(* IEC 61131-3 sources: Test-Git_ESME26/TestProgettoESME_26.fbsproj/PacDriveLib Migration/Motion/Positioning, 3 files *)

(* ---- PDL_FB_EndlessFeed.fb.st ---- *)
FUNCTION_BLOCK PDL_FB_EndlessFeed

VAR_INPUT
	i_xEnable					: BOOL;			(* Enable of FB *)
	i_ifDrive					: MOIN.IF_Axis;	(* Axis *)
	i_lrVel 					: LREAL;		(* Ceiling velocity in units/sec, -MaxVel to +MaxVel *)
	i_lrAcc  					: LREAL;		(* Acceleration units/s^2, value: 0...lrLimitMaxAccDec *)
	i_lrDec 					: LREAL;		(* Deceleration units/s^2, value: 0...lrLimitMaxAccDec *)
	i_lrJerk					: LREAL;		(* Jerk units/s^3, value: >0 *)
	i_lrPeriod					: LREAL;		(* LINEAR axis: the position is kept within the period value (0 … i_lrPeriod), in units, must be > 0
												   MODULO axis: value is ignored -> period is read from axis (i_ifDrive.lrModuloPeriod)  *)
	i_lrStopPosition			: LREAL;		(* 0 <= StopPosition <= Periode*)
	i_xStart					: BOOL;			(* starts with pos. edge *)
END_VAR

VAR_OUTPUT
	q_xActive					: BOOL;			(* FB enabled*)
	q_xReady					: BOOL;
	q_etDiag					: GD.ET_Diag := GD.ET_Diag.Ok;
	q_etDiagExt					: PDL_ET_DiagExt := PDL_ET_DiagExt.Disabled;
	q_sMsg						: STRING[80];
	q_xMotionInstructionActive	: BOOL;			(* axis is moving *)
	q_lrPosition				: LREAL;		(* axis position *)
	q_xInVelocity				: BOOL;			(* Velocity > VEL*0.99 AND Velocity < VEL* 1.01) *)
END_VAR

VAR
	xInterfacesInitialised		: BOOL;
	xEnableFlag					: BOOL;
	diState						: DINT;

	xMoveToStoppingStarted		: BOOL; //movement to lrStopPosition was started
	lrStopPosition				: LREAL;//calculated stopping position for linear axis when i_xStart = FALSE
	lrPeriodeCount				: LREAL;//periods needed for stopping
	lrStoppingDistance			: LREAL;//distance needed for stopping with actual vel, acc
	stStoppingDistance			: MOIN.ST_Trajectory;
	xErrorCalcStopping			: BOOL;
	etResultCalcStopping		: MOIN.ET_Result;

	//actual active values
	lrActVel					: LREAL;
	lrActJerk					: LREAL;
	lrAccel						: LREAL;
	lrDecel						: LREAL;

	fbLoggerPoint				: APL.FB_LoggerPoint;

	fbSetPos					: PLCO.MC_SetPosition;
	lrInchPos					: LREAL;

	fbStop						: PLCO.MC_Stop;
	fbMoveVelocity				: PLCO.MC_MoveVelocity;
	fbMoveAbsolute				: PLCO.MC_MoveAbsolute;
	fbHalt						: PLCO.MC_Halt;
	xExecuteHalt				: BOOL;

	xModuloAxis					: BOOL;
	lrModuloPeriod				: LREAL;

	xSuccess					: BOOL;
	ifGetParentDevice   		: DTSI.IF_GetParentDevice;
	ifDeviceAccess      		: DTSI.IF_DeviceAccess;
	ifDriveConfigAccess			: DDI.IF_DriveConfigAccess;
	ifDriveConfig				: DDI.IF_DriveConfig;

	ifDeviceTreeObjectAccess      : UFMPLCI.IF_DeviceTreeObjectAccess;
	sDriveName                    : STRING(80);

END_VAR

(*--------------------------------------------------------------------------------------------------------------------------------------------*)
//Enable
{region "enable"}
IF i_xEnable AND NOT xEnableFlag THEN

	xEnableFlag := TRUE;

	THIS^.fbLoggerPoint.AddLogEntry(	i_etLogLevel	:= APL.ET_LogLevel.UserAction,
										i_etDiag		:= q_etDiag,
										i_udiDiagExt	:= q_etDiagExt,
										i_sMessage		:= 'enable function block');

	xMoveToStoppingStarted 		:= FALSE;
	q_xActive					:= TRUE;
	q_xMotionInstructionActive	:= FALSE;
	q_xInVelocity				:= FALSE;
	q_xReady					:= FALSE;
	diState 					:= 0;

	SetDiagOutput(	i_etDiag	:= GD.ET_Diag.OK,
					i_etDiagExt := PDL_ET_DiagExt.Initializing,
					i_sMsg		:= '');

	xInterfacesInitialised := Init();
	IF NOT xInterfacesInitialised THEN
		RETURN;
	END_IF

	IF NOT InputParameterCheck() THEN
		RETURN;
	END_IF

	q_xReady := TRUE;
	lrActVel := 0;

	SetDiagOutput(	i_etDiag	:= GD.ET_Diag.OK,
					i_etDiagExt := PDL_ET_DiagExt.WaitForStart,
					i_sMsg		:= '');
	diState := 10;
{endregion}

(*--------------------------------------------------------------------------------------------------------------------------------------------*)
//Disable
{region "disable"}
ELSIF NOT i_xEnable AND xEnableFlag THEN
	xEnableFlag := FALSE;

	THIS^.fbLoggerPoint.AddLogEntry(	i_etLogLevel	:= APL.ET_LogLevel.UserAction,
										i_etDiag		:= q_etDiag,
										i_udiDiagExt	:= q_etDiagExt,
										i_sMessage		:= 'disable function block' );

	q_xInVelocity	:= FALSE;
	q_xReady		:= FALSE;

	IF xInterfacesInitialised THEN

		SetDiagOutput(	i_etDiag	:= GD.ET_Diag.OK,
						i_etDiagExt := PDL_ET_DiagExt.WaitUntilDisabled,
						i_sMsg		:= '');

		diState := 100;
	ELSE
		q_xActive					:= FALSE;
		q_xMotionInstructionActive	:= FALSE;
		q_lrPosition				:= 0.0;

		SetDiagOutput(	i_etDiag	:= GD.ET_Diag.OK,
						i_etDiagExt := PDL_ET_DiagExt.Disabled,
						i_sMsg		:= '');
		diState := 0;
	END_IF
END_IF
{endregion}

(*--------------------------------------------------------------------------------------------------------------------------------------------*)
// Cyclic when enabled
{region "cyclic"}
IF xInterfacesInitialised AND q_xActive THEN

	//restart after i_lrVel was 0
	IF    ABS(i_lrVel) > 0
	  AND diState = 30
	THEN
		xExecuteHalt := FALSE;
		THIS^.fbLoggerPoint.AddLogEntry(	i_etLogLevel	:= APL.ET_LogLevel.UserAction,
											i_etDiag		:= q_etDiag,
											i_udiDiagExt	:= q_etDiagExt,
											i_sMessage		:= Standard.CONCAT('start vel set: ', LREAL_TO_STRING(i_lrVel)), );
		IF xMoveToStoppingStarted THEN
			SetDiagOutput(	i_etDiag	:= GD.ET_Diag.OK,
							i_etDiagExt := PDL_ET_DiagExt.WaitUntilStopPositionReached,
							i_sMsg		:= '');
		END_IF
		q_xMotionInstructionActive	:= TRUE;
		diState := 10;
	END_IF

	//stop  (i_lrVel = 0)
	IF    (  i_xStart
		  OR q_xMotionInstructionActive
		  )
	  AND i_lrVel = 0
	  AND diState = 10
	THEN
		IF i_xStart THEN
			THIS^.fbLoggerPoint.AddLogEntry(	i_etLogLevel	:= APL.ET_LogLevel.UserAction,
												i_etDiag		:= q_etDiag,
												i_udiDiagExt	:= q_etDiagExt,
												i_sMessage		:= Standard.CONCAT('start with vel: ', LREAL_TO_STRING(i_lrVel)));
		ELSE
			THIS^.fbLoggerPoint.AddLogEntry(	i_etLogLevel	:= APL.ET_LogLevel.UserAction,
												i_etDiag		:= q_etDiag,
												i_udiDiagExt	:= q_etDiagExt,
												i_sMessage		:= Standard.CONCAT('stop vel set: ', LREAL_TO_STRING(i_lrVel)));
		END_IF

		SetDiagOutput(	i_etDiag	:= GD.ET_Diag.Ok,
						i_etDiagExt := PDL_ET_DiagExt.WaitForVelUnequalZero,
						i_sMsg		:= '');

		lrActVel := i_lrVel;
		xMoveToStoppingStarted := NOT i_xStart;
		q_xMotionInstructionActive	:= TRUE;
		xExecuteHalt := TRUE;
		diState := 30;
	END_IF

	//error
	IF  (	i_ifDrive.etAxisState = MOIN.ET_AxisState.ErrorStop
	  	OR  i_ifDrive.etAxisState = MOIN.ET_AxisState.Disabled
		)
		AND diState > 0
		AND diState < 100
	THEN
		diState := 0;

		q_xReady					:= FALSE;
		q_xMotionInstructionActive	:= FALSE;
		q_xInVelocity				:= FALSE;
		IF i_ifDrive.etAxisState = MOIN.ET_AxisState.Disabled THEN
			SetDiagOutput(	i_etDiag	:= GD.ET_Diag.DriveConditionInvalid,
							i_etDiagExt := PDL_ET_DiagExt.DriveNotReady,
							i_sMsg		:= STANDARD.CONCAT(sDriveName,' is DISABLED'));
		END_IF
		IF i_ifDrive.etAxisState = MOIN.ET_AxisState.ErrorStop THEN
			SetDiagOutput(	i_etDiag	:= GD.ET_Diag.DriveConditionInvalid,
							i_etDiagExt := PDL_ET_DiagExt.DriveNotReady,
							i_sMsg		:= STANDARD.CONCAT(sDriveName,' is ERRORSTOP'));
		END_IF
	END_IF

	//set q_lrPosition
	q_lrPosition	:= i_ifDrive.lrPosition;

	//linear axis only -> set new position when q_lrPosition > i_lrPeriod
	IF NOT xModuloAxis THEN
		SetPos();
	END_IF
END_IF
{endregion}

(*--------------------------------------------------------------------------------------------------------------------------------------------*)
// State machine
CASE  diState OF

(*********************************************************************************************************************)
	0:	//Error or Not Enabled
		;

(*********************************************************************************************************************)
	10: //endless movement and positioning to stop pos
{region "endlessMovementAndPositioning"}
		fbStop( Execute := FALSE );
		fbHalt( Execute := FALSE );

		fbMoveAbsolute( );
		fbMoveVelocity( );

		SetInVelocity();

		//wait for stop position reached
		IF fbMoveAbsolute.Done THEN
			fbMoveAbsolute( Execute := FALSE);
			xMoveToStoppingStarted := FALSE;

			q_xInVelocity				:= FALSE;
			q_xMotionInstructionActive	:= FALSE;

			SetDiagOutput(	i_etDiag	:= GD.ET_Diag.OK,
							i_etDiagExt := PDL_ET_DiagExt.WaitForStart,
							i_sMsg		:= '');
		END_IF

		//start movement to stopPosition...
		IF    NOT i_xStart  //...when input i_xStart is set to false
		  AND q_xMotionInstructionActive
		  AND NOT xMoveToStoppingStarted
		  OR  i_lrVel <> lrActVel  //... when velocity changed
		  AND xMoveToStoppingStarted
		  AND q_xMotionInstructionActive
		THEN
			IF NOT xMoveToStoppingStarted THEN
				fbLoggerPoint.AddLogEntry(	i_etLogLevel	:= APL.ET_LogLevel.UserAction,
											i_etDiag		:= q_etDiag,
											i_udiDiagExt	:= q_etDiagExt,
											i_sMessage		:= 'stop movement');
			ELSE
				fbLoggerPoint.AddLogEntry(	i_etLogLevel	:= APL.ET_LogLevel.DebugMessage,
											i_etDiag		:= q_etDiag,
											i_udiDiagExt	:= q_etDiagExt,
											i_sMessage		:= Standard.CONCAT('new vel set: ', LREAL_TO_STRING(i_lrVel)) );
			END_IF

			MoveToStopPosition(); //calculate position and call fb
			xMoveToStoppingStarted := TRUE;

		//start Endless movement...
		ELSIF    i_xStart //...when input i_xStart is set to true
			AND (   NOT q_xMotionInstructionActive
				OR  xMoveToStoppingStarted
				)
			OR  i_lrVel <> lrActVel //... when velocity changed
			AND q_xMotionInstructionActive
		THEN
			xMoveToStoppingStarted := FALSE;
			IF lrActVel <> 0 THEN
				fbLoggerPoint.AddLogEntry(	i_etLogLevel	:= APL.ET_LogLevel.UserAction,
											i_etDiag		:= q_etDiag,
											i_udiDiagExt	:= q_etDiagExt,
											i_sMessage		:= Standard.CONCAT('start with vel: ', LREAL_TO_STRING(i_lrVel)) );
			END_IF

			MoveVelocity();//call fb
		END_IF

		//error
		IF fbMoveAbsolute.Error THEN
			q_xMotionInstructionActive	:= FALSE;
			q_xInVelocity				:= FALSE;

			SetDiagOutput(	i_etDiag	:= GD.ET_Diag.UnexpectedProgramBehavior,
							i_etDiagExt := PDL_ET_DiagExt.UnexpectedFeedback,
							i_sMsg		:= CONCAT('MC_MoveAbsolute.ErrorID: ', PLCO.FC_EtResultToString(fbMoveAbsolute.ErrorID) ));
			diState := 100;
		END_IF

		IF fbMoveVelocity.Error THEN
			q_xMotionInstructionActive	:= FALSE;
			q_xInVelocity				:= FALSE;

			SetDiagOutput(	i_etDiag	:= GD.ET_Diag.UnexpectedProgramBehavior,
							i_etDiagExt := PDL_ET_DiagExt.UnexpectedFeedback,
							i_sMsg		:= CONCAT('MC_MoveVelocity.ErrorID: ', PLCO.FC_EtResultToString(fbMoveVelocity.ErrorID) ));
			diState := 100;
		END_IF
{endregion}

(*********************************************************************************************************************)
	30:	//stop  (i_lrVel = 0)
{region "stop (i_lrVel = 0)"}
		fbMoveAbsolute( Execute := FALSE );
		fbMoveVelocity( Execute := FALSE );
		fbStop( Execute := FALSE );

		fbHalt( Execute 		:= xExecuteHalt,
				Deceleration 	:= i_lrDec,
				Jerk			:= lrActJerk);

		q_xInVelocity := 	(  xMoveToStoppingStarted
							OR q_xMotionInstructionActive
							)
						AND NOT fbHalt.Active;

		//stopping done
		IF fbHalt.Done THEN
			xExecuteHalt := FALSE;
			IF xMoveToStoppingStarted THEN
				q_xMotionInstructionActive	:= FALSE;//only reset when stopping was started
			END_IF
		END_IF

		//restarted after stopping
		IF 	     i_xStart
			 AND xMoveToStoppingStarted
		THEN
			xMoveToStoppingStarted := FALSE;
			q_xMotionInstructionActive	:= TRUE;

		//vel was 0 and start is set to false
		ELSIF    NOT i_xStart
			 AND NOT xMoveToStoppingStarted
		THEN
			xExecuteHalt := FALSE;
			q_xInVelocity	:= FALSE;
			fbLoggerPoint.AddLogEntry(	i_etLogLevel	:= APL.ET_LogLevel.UserAction,
										i_etDiag		:= q_etDiag,
										i_udiDiagExt	:= q_etDiagExt,
										i_sMessage		:= 'stop movement');
			SetDiagOutput(	i_etDiag	:= GD.ET_Diag.OK,
							i_etDiagExt := PDL_ET_DiagExt.WaitForStart,
							i_sMsg		:= '');
			q_xMotionInstructionActive	:= FALSE;
			diState := 10;
		END_IF

		//error
		IF fbHalt.Error THEN
			q_xMotionInstructionActive	:= FALSE;
			q_xInVelocity				:= FALSE;
			xExecuteHalt				:= FALSE;

			SetDiagOutput(	i_etDiag	:= GD.ET_Diag.UnexpectedProgramBehavior,
							i_etDiagExt := PDL_ET_DiagExt.UnexpectedFeedback,
							i_sMsg		:= CONCAT('MC_Halt.ErrorID: ', PLCO.FC_EtResultToString(fbHalt.ErrorID) ));
			diState := 100;
		END_IF
{endregion}

(*********************************************************************************************************************)
	100: //controller stop
{region "controllerStop"}
		fbMoveAbsolute( Execute := FALSE );
		fbMoveVelocity( Execute := FALSE );
		fbHalt( Execute := FALSE );

		IF 	  i_ifDrive.etAxisState <> MOIN.ET_AxisState.Disabled
		  AND i_ifDrive.etAxisState <> MOIN.ET_AxisState.ErrorStop
		  AND i_ifDrive.etAxisState <> MOIN.ET_AxisState.Standstill
		  AND i_ifDrive.etAxisState <> MOIN.ET_AxisState.Stopping
		THEN
			fbStop.Execute 			:= TRUE;
			fbStop.Deceleration 	:= i_ifDrive.lrErrorStopDec;
			fbStop.Jerk 			:= i_ifDrive.lrErrorStopJerk;
		END_IF

		fbStop();

		//stopping done
		IF 	  i_ifDrive.etAxisState = MOIN.ET_AxisState.Disabled
		  OR  i_ifDrive.etAxisState = MOIN.ET_AxisState.ErrorStop
		  OR  i_ifDrive.etAxisState = MOIN.ET_AxisState.Standstill
		  OR  fbStop.Done
		THEN
			q_xMotionInstructionActive	:= FALSE;
			q_xReady := FALSE;
			fbStop( Execute := FALSE );

			IF NOT i_xEnable THEN
				xInterfacesInitialised := FALSE;

				q_xMotionInstructionActive	:= FALSE;
				q_xActive					:= FALSE;

				SetDiagOutput(	i_etDiag	:= GD.ET_Diag.OK,
								i_etDiagExt := PDL_ET_DiagExt.Disabled,
								i_sMsg		:= '');
			END_IF

			diState := 0;
		END_IF

		//error
		IF fbStop.Error AND fbStop.ErrorId <> PLCO.ET_Result.StoppingInterrupted THEN
			q_xMotionInstructionActive	:= FALSE;
			q_xInVelocity				:= FALSE;

			SetDiagOutput(	i_etDiag	:= GD.ET_Diag.UnexpectedProgramBehavior,
							i_etDiagExt := PDL_ET_DiagExt.UnexpectedFeedback,
							i_sMsg		:= CONCAT('MC_Stop.ErrorID: ', PLCO.FC_EtResultToString(fbStop.ErrorID) ));
			fbStop( Execute := FALSE );
		END_IF
{endregion}

END_CASE
(*--------------------------------------------------------------------------------------------------------------------------------------------*)

(* ---- PDL_FB_Jogging.fb.st ---- *)
FUNCTION_BLOCK PDL_FB_Jogging
VAR_INPUT
	i_xEnable					: BOOL;				(* enables the FB *)
	i_ifDrive					: MOIN.IF_Axis;		(* Axis *)
	i_xJogForw					: BOOL;				(* Jogging Forward *)
	i_xJogBack					: BOOL;				(* Jogging Backward *)
	i_lrPeriod					: LREAL;			(* if Periode = 0 --> no Position manipulation *)
	i_xEndless					: BOOL;				(* TRUE = jogging endless, FALSE = jogging with max Distance of Step *)
	i_lrMaxDistance				: LREAL;			(* Step  in Units *)
	i_lrVel						: LREAL;			(* ceiling velocity in U/sec; 0<=Vel<Velmax*)
	i_lrAcc						: LREAL;			(* Acceleration units/s^2, value: 0...lrLimitMaxAccDec *)
	i_lrDec						: LREAL;			(* Deceleration units/s^2, value: 0...lrLimitMaxAccDec *)
	i_lrJerk					: LREAL;
END_VAR

VAR_OUTPUT
	q_xActive					: BOOL;				(* TRUE if  FB is enabled *)
	q_xReady					: BOOL;
	q_etDiag					: GD.ET_Diag := GD.ET_Diag.Ok;
	q_etDiagExt					: PDL_ET_DiagExt := PDL_ET_DiagExt.Disabled;
	q_sMsg						: STRING[80];
	q_xMotionInstructionActive	: BOOL;				(* TRUE if motion is active *)
	q_lrPosition				: LREAL;			(* shows the Reference position of the axis *)
	q_xStepFinished				: BOOL;				(* TRUE if step is done *)
END_VAR

VAR
	xInterfacesInitialised		: BOOL;
	fbLoggerPoint				: APL.FB_LoggerPoint;

	diState						: DINT;
	xEnableFlag					: BOOL;
	iPeriodeCount				: INT;
	lrPosBuffer					: LREAL;

	fbSetPos					: PLCO.MC_SetPosition;
	fbStop						: PLCO.MC_Stop;
	fbJog						: PLCO.MC_Jog;
	xJogForwardStarted			: BOOL; //FALSE: jogging backward, TRUE: jogging forward,

	xSuccess					: BOOL;
	ifGetParentDevice   		: DTSI.IF_GetParentDevice;
	ifDeviceAccess      		: DTSI.IF_DeviceAccess;
	ifDriveConfigAccess			: DDI.IF_DriveConfigAccess;
	ifDriveConfig				: DDI.IF_DriveConfig;

	ifDeviceTreeObjectAccess      : UFMPLCI.IF_DeviceTreeObjectAccess;
	sDriveName                    : STRING(80);

END_VAR

(*--------------------------------------------------------------------------------------------------------------------------------------------*)
//Enable
{region "enable"}
IF i_xEnable AND NOT xEnableFlag THEN
	xEnableFlag := TRUE;
	q_xActive					:= TRUE;
	q_xReady					:= FALSE;
	q_xMotionInstructionActive	:= FALSE;
	q_xStepFinished				:= FALSE;
	diState := 0;
	fbLoggerPoint.AddLogEntry(	i_etLogLevel	:= APL.ET_LogLevel.UserAction,
								i_etDiag		:= q_etDiag,
								i_udiDiagExt	:= q_etDiagExt,
								i_sMessage		:= 'enable function block');
	SetDiagOutput(	i_etDiag	:= GD.ET_Diag.OK,
					i_etDiagExt := PDL_ET_DiagExt.Initializing,
					i_sMsg		:= '');

	xInterfacesInitialised := Init();
	IF NOT xInterfacesInitialised THEN
		RETURN;
	END_IF

	IF NOT InputParameterCheck( xCheckDistance := FALSE, xCheckPeriod := FALSE ) THEN
		RETURN;
	END_IF

	//check axis state
	IF  (	i_ifDrive.etAxisState = MOIN.ET_AxisState.ErrorStop
	  	OR  i_ifDrive.etAxisState = MOIN.ET_AxisState.Disabled
		)
	THEN
		IF i_ifDrive.etAxisState = MOIN.ET_AxisState.Disabled THEN
			SetDiagOutput(	i_etDiag	:= GD.ET_Diag.DriveConditionInvalid,
							i_etDiagExt := PDL_ET_DiagExt.DriveNotReady,
							i_sMsg		:= STANDARD.CONCAT(sDriveName,' is DISABLED'));
		END_IF
		IF i_ifDrive.etAxisState = MOIN.ET_AxisState.ErrorStop THEN
			SetDiagOutput(	i_etDiag	:= GD.ET_Diag.DriveConditionInvalid,
							i_etDiagExt := PDL_ET_DiagExt.DriveNotReady,
							i_sMsg		:= STANDARD.CONCAT(sDriveName,' is ERRORSTOP'));
		END_IF

	ELSE
		//set q_lrPosition
		IF NOT SetPos() THEN
			RETURN;
		END_IF
		q_xReady := TRUE;
		SetDiagOutput(	i_etDiag	:= GD.ET_Diag.Ok,
						i_etDiagExt := PDL_ET_DiagExt.WaitForJoggingInputsLow,
						i_sMsg		:= '');

		fbJog(	JogForward := FALSE, JogBackward := FALSE );
		fbStop( Execute := FALSE );
		diState := 10;
	END_IF
{endregion}

(*--------------------------------------------------------------------------------------------------------------------------------------------*)
//Disable
{region "disable"}
ELSIF NOT i_xEnable AND xEnableFlag THEN
	xEnableFlag := FALSE;
	fbLoggerPoint.AddLogEntry(	i_etLogLevel	:= APL.ET_LogLevel.UserAction,
								i_etDiag		:= q_etDiag,
								i_udiDiagExt	:= q_etDiagExt,
								i_sMessage		:= 'disable function block');
	q_xReady		:= FALSE;
	q_xStepFinished	:= FALSE;
	IF xInterfacesInitialised THEN
		SetDiagOutput(	i_etDiag	:= GD.ET_Diag.Ok,
						i_etDiagExt := PDL_ET_DiagExt.WaitUntilDisabled,
						i_sMsg		:= '');
		diState := 100;
	ELSE
		q_xActive					:= FALSE;
		q_xMotionInstructionActive	:= FALSE;
		q_lrPosition				:= 0.0;
		SetDiagOutput(	i_etDiag	:= GD.ET_Diag.Ok,
						i_etDiagExt := PDL_ET_DiagExt.Disabled,
						i_sMsg		:= '');
		diState := 0;
	END_IF
END_IF
{endregion}

(*--------------------------------------------------------------------------------------------------------------------------------------------*)
// Cyclic when enabled
{region "cyclic"}
IF xInterfacesInitialised AND q_xActive THEN

	//error
	IF  (	i_ifDrive.etAxisState = MOIN.ET_AxisState.ErrorStop
	  	OR  i_ifDrive.etAxisState = MOIN.ET_AxisState.Disabled
		)
		AND diState > 0
		AND diState < 100
	THEN
		diState := 0;

		q_xReady					:= FALSE;
		q_xStepFinished				:= FALSE;
		q_xMotionInstructionActive	:= FALSE;

		IF i_ifDrive.etAxisState = MOIN.ET_AxisState.Disabled THEN
			SetDiagOutput(	i_etDiag	:= GD.ET_Diag.DriveConditionInvalid,
							i_etDiagExt := PDL_ET_DiagExt.DriveNotReady,
							i_sMsg		:= ' Axis is DISABLED');
		END_IF
		IF i_ifDrive.etAxisState = MOIN.ET_AxisState.ErrorStop THEN
			SetDiagOutput(	i_etDiag	:= GD.ET_Diag.DriveConditionInvalid,
							i_etDiagExt := PDL_ET_DiagExt.DriveNotReady,
							i_sMsg		:= ' Axis in ERRORSTOP');
		END_IF
	END_IF

	//set q_lrPosition
	SetPos();

END_IF
{endregion}

(*--------------------------------------------------------------------------------------------------------------------------------------------*)
// State machine
CASE  diState OF

(*********************************************************************************************************************)
	0://Error or Not Enabled
		;

(*********************************************************************************************************************)
	10:	// Wait for jogging inputs low
{region "wait for inputs reset"}
		IF NOT i_xJogForw AND NOT i_xJogBack THEN
			SetDiagOutput(	i_etDiag	:= GD.ET_Diag.Ok,
							i_etDiagExt := PDL_ET_DiagExt.WaitForJogging,
							i_sMsg		:= '');
			diState := 20;
		END_IF
{endregion}

(*********************************************************************************************************************)
	20:	//Wait for start
{region "wait for start"}
		IF i_xJogForw OR i_xJogBack THEN
			xJogForwardStarted := i_xJogForw;

			//set logger msg
			IF i_xJogForw THEN
				fbLoggerPoint.AddLogEntry(	i_etLogLevel	:= APL.ET_LogLevel.UserAction,
											i_etDiag		:= q_etDiag,
											i_udiDiagExt	:= q_etDiagExt,
											i_sMessage		:= 'Jog Forward' );
			ELSE
				fbLoggerPoint.AddLogEntry(	i_etLogLevel	:= APL.ET_LogLevel.UserAction,
											i_etDiag		:= q_etDiag,
											i_udiDiagExt	:= q_etDiagExt,
											i_sMessage		:= 'Jog Backward' );
			END_IF

			//check inputs
			IF NOT InputParameterCheck() THEN
				q_xReady := FALSE;
				diState  := 0;

			ELSE
				//start movement
				IF i_xEndless THEN
					fbJog.JogType := PLCO.MC_JogType.Velocity;
				ELSE
					fbJog.JogType := PLCO.MC_JogType.PositionOffset;
				END_IF

				fbJog(	JogForward		:= i_xJogForw,
						JogBackward		:= i_xJogBack AND NOT i_xJogForw, //if both inputs are true -> move forward
						Position		:= i_lrMaxDistance,
						Velocity		:= i_lrVel,
						Acceleration	:= i_lrAcc,
						Deceleration	:= i_lrDec,
						Jerk			:= i_lrJerk );

				IF fbJog.Error THEN
					diState:= 0;
					q_xMotionInstructionActive	:= FALSE;
					SetDiagOutput(	i_etDiag	:= GD.ET_Diag.UnexpectedProgramBehavior,
									i_etDiagExt := PDL_ET_DiagExt.UnexpectedFeedback,
									i_sMsg		:= CONCAT('MC_Jog.ErrorId: ', TO_STRING(fbJog.ErrorId)));
					fbJog( JogForward := FALSE, JogBackward := FALSE );
					RETURN;
				END_IF

				q_xMotionInstructionActive	:= TRUE;
				q_xStepFinished				:= FALSE;

				//set diag output
				IF i_xJogForw THEN
					SetDiagOutput(	i_etDiag	:= GD.ET_Diag.Ok,
									i_etDiagExt := PDL_ET_DiagExt.JoggingForward,
									i_sMsg		:= '');
				ELSE
					SetDiagOutput(	i_etDiag	:= GD.ET_Diag.Ok,
									i_etDiagExt := PDL_ET_DiagExt.JoggingBackward,
									i_sMsg		:= '');
				END_IF

				diState := 30;
			END_IF
		END_IF
{endregion}

(*********************************************************************************************************************)
	30:	//jogging movement active
{region "jogging active"}
		fbJog();

		//stop jogging movement
		IF    fbJog.Busy
		  AND (   NOT i_xJogForw AND xJogForwardStarted
		      OR  NOT i_xJogBack AND NOT xJogForwardStarted
			  )
		THEN
			IF xJogForwardStarted THEN
				fbLoggerPoint.AddLogEntry(	i_etLogLevel	:= APL.ET_LogLevel.UserAction,
											i_etDiag		:= q_etDiag,
											i_udiDiagExt	:= q_etDiagExt,
											i_sMessage		:= 'Hold jogging forward');
			ELSE
				fbLoggerPoint.AddLogEntry(	i_etLogLevel	:= APL.ET_LogLevel.UserAction,
											i_etDiag		:= q_etDiag,
											i_udiDiagExt	:= q_etDiagExt,
											i_sMessage		:= 'Hold jogging backward');
			END_IF

			fbJog(	JogForward := FALSE, JogBackward := FALSE );

			SetDiagOutput(	i_etDiag	:= GD.ET_Diag.Ok,
							i_etDiagExt := PDL_ET_DiagExt.WaitUntilStopped,
							i_sMsg		:= '');
			diState := 50;

		//target pos reached: go to waiting step when inputs are false
		ELSIF fbJog.Done AND NOT i_xJogForw AND NOT i_xJogBack THEN
			fbJog(	JogForward := FALSE, JogBackward := FALSE );

			IF xJogForwardStarted THEN
				fbLoggerPoint.AddLogEntry(	i_etLogLevel	:= APL.ET_LogLevel.UserAction,
											i_etDiag		:= q_etDiag,
											i_udiDiagExt	:= q_etDiagExt,
											i_sMessage		:= 'Finished jogging forward');
			ELSE
				fbLoggerPoint.AddLogEntry(	i_etLogLevel	:= APL.ET_LogLevel.UserAction,
											i_etDiag		:= q_etDiag,
											i_udiDiagExt	:= q_etDiagExt,
											i_sMessage		:= 'Finished jogging backward');
			END_IF
			q_xMotionInstructionActive	:= FALSE;
			q_xStepFinished				:= TRUE;

			SetDiagOutput(	i_etDiag	:= GD.ET_Diag.Ok,
							i_etDiagExt := PDL_ET_DiagExt.WaitForJogging,
							i_sMsg		:= '');
			diState := 20;

		//target pos reached: set diag mesg
		ELSIF fbJog.Done THEN
			IF NOT q_xStepFinished THEN
				fbLoggerPoint.AddLogEntry(	i_etLogLevel	:= APL.ET_LogLevel.StatusMessage,
											i_etDiag		:= q_etDiag,
											i_udiDiagExt	:= q_etDiagExt,
											i_sMessage		:= 'Jog target reached',
											q_etDiag		=> ,
											q_etDiagExt		=> );
			END_IF
			q_xMotionInstructionActive	:= FALSE;
			q_xStepFinished				:= TRUE;
		END_IF

		//error
		IF fbJog.Error THEN
			q_xMotionInstructionActive	:= FALSE;
			q_xStepFinished				:= FALSE;
			q_xReady					:= FALSE;
			SetDiagOutput(	i_etDiag	:= GD.ET_Diag.UnexpectedProgramBehavior,
							i_etDiagExt := PDL_ET_DiagExt.UnexpectedFeedback,
							i_sMsg		:= CONCAT('MC_Jog.ErrorId: ', TO_STRING(fbJog.ErrorId)));
			fbJog( JogForward := FALSE, JogBackward := FALSE );
			diState := 0;
		END_IF
{endregion}

(*********************************************************************************************************************)
	50://wait for jogging movement stopped
{region "waitForJoggingMovementStopped"}
		fbJog(	JogForward := FALSE, JogBackward := FALSE );

		IF i_ifDrive.etAxisState = MOIN.ET_AxisState.Standstill THEN
			q_xMotionInstructionActive	:= FALSE;
			SetDiagOutput(	i_etDiag	:= GD.ET_Diag.Ok,
							i_etDiagExt := PDL_ET_DiagExt.WaitForJogging,
							i_sMsg		:= '');
			diState := 20;

		ELSIF i_xJogForw OR i_xJogBack THEN
			diState := 20;
		END_IF
{endregion}

(*********************************************************************************************************************)
	100: //controller stop
{region "controllerstop"}
		fbJog(	JogForward := FALSE, JogBackward := FALSE );

		IF 	  i_ifDrive.etAxisState <> MOIN.ET_AxisState.Disabled
		  AND i_ifDrive.etAxisState <> MOIN.ET_AxisState.ErrorStop
		  AND i_ifDrive.etAxisState <> MOIN.ET_AxisState.Standstill
		  AND i_ifDrive.etAxisState <> MOIN.ET_AxisState.Stopping
		THEN
			fbStop.Execute 			:= TRUE;
			fbStop.Deceleration 	:= i_ifDrive.lrErrorStopDec;
			fbStop.Jerk 			:= i_ifDrive.lrErrorStopJerk;
		END_IF

		fbStop();

		//stopping done
		IF 	  i_ifDrive.etAxisState = MOIN.ET_AxisState.Disabled
		  OR  i_ifDrive.etAxisState = MOIN.ET_AxisState.ErrorStop
		  OR  i_ifDrive.etAxisState = MOIN.ET_AxisState.Standstill
		  OR  fbStop.Done
		THEN
			xInterfacesInitialised := FALSE;
			q_xMotionInstructionActive	:= FALSE;
			q_xStepFinished				:= FALSE;
			q_xActive					:= FALSE;
			q_xReady					:= FALSE;
			q_lrPosition				:= 0.0;
			fbStop( Execute := FALSE );

			SetDiagOutput(	i_etDiag	:= GD.ET_Diag.OK,
							i_etDiagExt := PDL_ET_DiagExt.Disabled,
							i_sMsg		:= '');

			diState := 0;
		END_IF

		//error
		IF fbStop.Error AND fbStop.ErrorId <> PLCO.ET_Result.StoppingInterrupted THEN
			q_xMotionInstructionActive	:= FALSE;

			SetDiagOutput(	i_etDiag	:= GD.ET_Diag.UnexpectedProgramBehavior,
							i_etDiagExt := PDL_ET_DiagExt.UnexpectedFeedback,
							i_sMsg		:= CONCAT('MC_Stop.ErrorID: ', PLCO.FC_EtResultToString(fbStop.ErrorID) ));
			fbStop( Execute := FALSE );
		END_IF
{endregion}

END_CASE
(*--------------------------------------------------------------------------------------------------------------------------------------------*)

(* ---- PDL_FB_VarioPosJerk.fb.st ---- *)
FUNCTION_BLOCK PDL_FB_VarioPosJerk

VAR_INPUT
	i_xEnable					: BOOL;				(* Enable of FB *)
	i_ifDrive					: MOIN.IF_Axis; 	(* Axis *)
	i_xStart					: BOOL;				(* Starts with pos. edge *)
	i_xStop						: BOOL;				(* Stops with pos. level *)
	i_lrTarget  				: LREAL;			(* target position or distance in [U] *)
	i_lrVel						: LREAL;			(* ceiling velocity in U/sec *)
	i_lrAcc						: LREAL;			(* Acceleration units/s^2, value: 0...lrLimitMaxAccDec *)
	i_lrDec						: LREAL;			(* Deceleration units/s^2, value: 0...lrLimitMaxAccDec *)
	i_lrJerk					: LREAL;			(* Jerk units/s^3, value: >0 *)
	i_etPosMode					: PDL_ET_PosMode;	(* POS_ENDLESS, POS_RELATIVE, POS_ABSOLUTE *)
END_VAR

VAR_OUTPUT
	q_xActive					: BOOL;				(* FB enabled *)
	q_xReady					: BOOL;
	q_etDiag					: GD.ET_Diag := GD.ET_Diag.OK;
	q_etDiagExt					: PDL_ET_DiagExt := PDL_ET_DiagExt.Disabled;
	q_sMsg						: STRING[80];
	q_xMotionInstructionActive	: BOOL;				(* axis is moving *)
	q_lrPosition				: LREAL;			(* axis position *)
	q_xInPosition				: BOOL;				(* target position reached *)
END_VAR

VAR
	xInterfacesInitialised		: BOOL;

	xEnableFlag					: BOOL;
	diState						: DINT;
	fbRtrigStartEdge			: Standard.R_TRIG;
	lrTarget					: LREAL; //for setting diag msg
	etActivePosMode				: PDL_ET_PosMode;

	fbLoggerPoint				: APL.FB_LoggerPoint;

	fbHalt						: PLCO.MC_Halt;
	fbStop						: PLCO.MC_Stop;
	fbMoveAbsolute				: PLCO.MC_MoveAbsolute;
	fbMoveRelative				: PLCO.MC_MoveRelative;
	fbSetPos					: PLCO.MC_SetPosition;

	xSuccess					: BOOL;
	ifGetParentDevice   		: DTSI.IF_GetParentDevice;
	ifDeviceAccess      		: DTSI.IF_DeviceAccess;
	ifDriveConfigAccess			: DDI.IF_DriveConfigAccess;
	ifDriveConfig				: DDI.IF_DriveConfig;

	ifDeviceTreeObjectAccess      : UFMPLCI.IF_DeviceTreeObjectAccess;
	sDriveName                    : STRING(80);

END_VAR

(*--------------------------------------------------------------------------------------------------------------------------------------------*)
//Enable
{region "enable"}
IF i_xEnable AND NOT xEnableFlag THEN
	xEnableFlag := TRUE;
	fbLoggerPoint.AddLogEntry(	i_etLogLevel	:= APL.ET_LogLevel.UserAction,
								i_etDiag		:= q_etDiag,
								i_udiDiagExt	:= q_etDiagExt,
								i_sMessage		:= 'enable function block');

	q_xMotionInstructionActive	:= FALSE;
	q_xInPosition				:= FALSE;
	q_xActive					:= TRUE;
	q_xReady					:= FALSE;
	diState := 0;
	SetDiagOutput(	i_etDiag	:= GD.ET_Diag.OK,
					i_etDiagExt := PDL_ET_DiagExt.Initializing,
					i_sMsg		:= '');

	xInterfacesInitialised := Init();
	IF NOT xInterfacesInitialised THEN
		RETURN;
	END_IF

	q_xReady := TRUE;
	SetDiagOutput(	i_etDiag	:= GD.ET_Diag.OK,
					i_etDiagExt := PDL_ET_DiagExt.WaitForStart,
					i_sMsg		:= '');
	diState	:= 10;
{endregion}

(*--------------------------------------------------------------------------------------------------------------------------------------------*)
//Disable
{region "disable"}
ELSIF NOT i_xEnable AND xEnableFlag THEN
	xEnableFlag := FALSE;
	fbLoggerPoint.AddLogEntry(	i_etLogLevel	:= APL.ET_LogLevel.UserAction,
								i_etDiag		:= q_etDiag,
								i_udiDiagExt	:= q_etDiagExt,
								i_sMessage		:= 'disable function block');

	IF xInterfacesInitialised THEN

		q_xMotionInstructionActive	:= FALSE;
		q_xInPosition				:= FALSE;
		q_xReady 					:= FALSE;

		SetDiagOutput(	i_etDiag	:= GD.ET_Diag.OK,
						i_etDiagExt := PDL_ET_DiagExt.WaitUntilDisabled,
						i_sMsg		:= '');

		diState						:= 100;
	ELSE
		q_xActive					:= FALSE;
		q_xReady					:= FALSE;
		q_xMotionInstructionActive	:= FALSE;
		q_xInPosition				:= FALSE;
		q_lrPosition				:= 0.0;
		SetDiagOutput(	i_etDiag	:= GD.ET_Diag.OK,
						i_etDiagExt := PDL_ET_DiagExt.Disabled,
						i_sMsg		:= '');
		diState := 0;
	END_IF
END_IF
{endregion}

(*--------------------------------------------------------------------------------------------------------------------------------------------*)
// Cyclic when enabled
{region "cyclic"}
IF xInterfacesInitialised AND q_xActive THEN

	//stop
	IF    i_xStop
	  AND q_xMotionInstructionActive
	  AND diState = 10 //positioning active
	THEN
		fbLoggerPoint.AddLogEntry(	i_etLogLevel	:= APL.ET_LogLevel.UserAction,
									i_etDiag		:= q_etDiag,
									i_udiDiagExt	:= q_etDiagExt,
									i_sMessage		:= 'stop positioning');

		SetDiagOutput(	i_etDiag	:= GD.ET_Diag.OK,
						i_etDiagExt := PDL_ET_DiagExt.Stopping,
						i_sMsg		:= '');

		diState := 30;
	END_IF

	//error
	IF  (	i_ifDrive.etAxisState = MOIN.ET_AxisState.ErrorStop
	  	OR  i_ifDrive.etAxisState = MOIN.ET_AxisState.Disabled
		)
		AND diState > 0
		AND diState < 100
	THEN
		q_xReady					:= FALSE;
		q_xMotionInstructionActive	:= FALSE;
		IF i_ifDrive.etAxisState = MOIN.ET_AxisState.Disabled THEN
			SetDiagOutput(	i_etDiag	:= GD.ET_Diag.DriveConditionInvalid,
							i_etDiagExt := PDL_ET_DiagExt.DriveNotReady,
							i_sMsg		:= STANDARD.CONCAT(sDriveName,' is DISABLED'));
		END_IF
		IF i_ifDrive.etAxisState = MOIN.ET_AxisState.ErrorStop THEN
			SetDiagOutput(	i_etDiag	:= GD.ET_Diag.DriveConditionInvalid,
							i_etDiagExt := PDL_ET_DiagExt.DriveNotReady,
							i_sMsg		:= STANDARD.CONCAT(sDriveName,' is ERRORSTOP'));
		END_IF
		diState := 0;
	END_IF

	q_lrPosition := i_ifDrive.lrPosition;
END_IF

fbRtrigStartEdge(CLK := i_xStart);
{endregion}

(*--------------------------------------------------------------------------------------------------------------------------------------------*)
// State machine
CASE  diState OF
(*********************************************************************************************************************)
	0: //Error or Not Enabled
		;

(*********************************************************************************************************************)
	10:	//positioning
{region "positioniong"}
		fbMoveAbsolute( Execute :=    q_xMotionInstructionActive
								  AND (	 etActivePosMode = PDL_ET_PosMode.Absolute
								  	  OR etActivePosMode = PDL_ET_PosMode.Endless
									  )
						);
		fbMoveRelative( Execute :=    q_xMotionInstructionActive
								  AND etActivePosMode = PDL_ET_PosMode.Relative
						);

		fbStop( Execute := FALSE );
		fbHalt( Execute := FALSE );

		// Wait for pos. edge of Start
		IF fbRtrigStartEdge.Q  AND NOT i_xStop THEN

			IF q_xMotionInstructionActive THEN
				fbLoggerPoint.AddLogEntry(	i_etLogLevel	:= APL.ET_LogLevel.UserAction,
											i_etDiag		:= q_etDiag,
											i_udiDiagExt	:= q_etDiagExt,
											i_sMessage		:= 'start new positioning');
			ELSE
				fbLoggerPoint.AddLogEntry(	i_etLogLevel	:= APL.ET_LogLevel.UserAction,
											i_etDiag		:= q_etDiag,
											i_udiDiagExt	:= q_etDiagExt,
											i_sMessage		:= 'start positioning');
			END_IF

			// error during parametercheck - diag output already set in method InputParameterCheck
			IF NOT InputParameterCheck() THEN
				q_xReady := FALSE;
				diState := 0;
				RETURN;
			END_IF

			q_xMotionInstructionActive	:= TRUE;
			q_xInPosition	:= FALSE;
			etActivePosMode	:= i_etPosMode;

			//execute  cmd
			SetPos();
			fbMoveAbsolute( Execute := FALSE );
			fbMoveRelative( Execute := FALSE );

			IF   i_etPosMode = PDL_ET_PosMode.Absolute
			  OR i_etPosMode = PDL_ET_PosMode.Endless
			THEN
				IF 	  (i_etPosMode = PDL_ET_PosMode.Endless  AND i_lrTarget >= 0)
				  OR  (i_etPosMode = PDL_ET_PosMode.Absolute AND (i_lrTarget - q_lrPosition) >= 0)
				THEN
					fbMoveAbsolute.Direction := MOIN.ET_Direction.PositiveDirection;
				ELSE
					fbMoveAbsolute.Direction := MOIN.ET_Direction.NegativeDirection;
				END_IF
				fbMoveAbsolute.Acceleration 	:= i_lrAcc;
				fbMoveAbsolute.Deceleration 	:= i_lrDec;
				fbMoveAbsolute.Velocity 		:= i_lrVel;
				fbMoveAbsolute.Jerk 			:= i_lrJerk;
				fbMoveAbsolute.Position			:= i_lrTarget;
				fbMoveAbsolute( Execute := TRUE );
			ELSE
				fbMoveRelative.Acceleration 	:= i_lrAcc;
				fbMoveRelative.Deceleration 	:= i_lrDec;
				fbMoveRelative.Velocity 		:= i_lrVel;
				fbMoveRelative.Jerk 			:= i_lrJerk;
				fbMoveRelative.Distance			:= i_lrTarget;
				fbMoveRelative( Execute := TRUE );
			END_IF

			//set diag msg
			IF    (i_etPosMode = PDL_ET_PosMode.Absolute)
			  OR  (i_etPosMode = PDL_ET_PosMode.Endless)
			THEN
				lrTarget := i_lrTarget;
			ELSIF (i_etPosMode = PDL_ET_PosMode.Relative) THEN
				lrTarget := i_lrTarget + i_ifDrive.lrPosition;
			END_IF
			SetDiagOutput(	i_etDiag	:= GD.ET_Diag.OK,
							i_etDiagExt := PDL_ET_DiagExt.Positioning,
							i_sMsg		:= SE_CTBX.FC_MultiConcat(	i_sString1	:= 'Mode: ',
																	i_sString2	:= etPosModeToString(i_etPosMode := i_etPosMode),
																	i_sString3	:= ' Target: ',
																	i_sString4	:= TO_STRING(i_lrTarget)) );
		//finished
		ELSIF    fbMoveAbsolute.Done
			 AND (	etActivePosMode = PDL_ET_PosMode.Absolute
				 OR etActivePosMode = PDL_ET_PosMode.Endless
				 )
			 OR  fbMoveRelative.Done
			 AND etActivePosMode = PDL_ET_PosMode.Relative
		THEN
			q_xMotionInstructionActive	:= FALSE;
			q_xInPosition	:= TRUE;
			SetDiagOutput(	i_etDiag	:= GD.ET_Diag.OK,
							i_etDiagExt := PDL_ET_DiagExt.WaitForStart,
							i_sMsg		:= '');
		END_IF

		//error
		IF fbMoveRelative.Error THEN
			q_xMotionInstructionActive	:= FALSE;

			SetDiagOutput(	i_etDiag	:= GD.ET_Diag.UnexpectedProgramBehavior,
							i_etDiagExt := PDL_ET_DiagExt.UnexpectedFeedback,
							i_sMsg		:= CONCAT('MC_MoveRelative.ErrorID: ', PLCO.FC_EtResultToString( fbMoveRelative.ErrorID ) ));
			diState	:= 100;
		END_IF

		IF fbMoveAbsolute.Error THEN
			q_xMotionInstructionActive	:= FALSE;

			SetDiagOutput(	i_etDiag	:= GD.ET_Diag.UnexpectedProgramBehavior,
							i_etDiagExt := PDL_ET_DiagExt.UnexpectedFeedback,
							i_sMsg		:= CONCAT('MC_MoveAbsolute.ErrorID: ', PLCO.FC_EtResultToString( fbMoveAbsolute.ErrorID ) ));
			diState	:= 100;
		END_IF
{endregion}

(*********************************************************************************************************************)
	30: //stop
{region "stop"}
       	fbMoveAbsolute( Execute := FALSE  );
       	fbMoveRelative( Execute := FALSE  );
		fbStop(  Execute := FALSE );

		fbHalt( Execute 		:= TRUE,
				Deceleration 	:= i_lrDec,
				Jerk 			:= i_lrJerk
				);

		//stopping done
		IF		fbHalt.Done
			OR  i_ifDrive.etAxisState = MOIN.ET_AxisState.Standstill
		THEN
			q_xMotionInstructionActive := FALSE;

			fbHalt(  Execute := FALSE );

			SetDiagOutput(	i_etDiag	:= GD.ET_Diag.OK,
							i_etDiagExt := PDL_ET_DiagExt.WaitForStart,
							i_sMsg		:= '');

			diState	:= 10;
		END_IF

		//error
		IF fbHalt.Error THEN
			q_xMotionInstructionActive	:= FALSE;

			SetDiagOutput(	i_etDiag	:= GD.ET_Diag.UnexpectedProgramBehavior,
							i_etDiagExt := PDL_ET_DiagExt.UnexpectedFeedback,
							i_sMsg		:= CONCAT('MC_Halt.ErrorID: ', PLCO.FC_EtResultToString( fbHalt.ErrorID ) ));
			diState	:= 100;
		END_IF
{endregion}

(*********************************************************************************************************************)
	100: //controller stop
{region "controllerStop"}
       	fbMoveAbsolute( Execute := FALSE  );
       	fbMoveRelative( Execute := FALSE  );
		fbHalt( Execute := FALSE );

		IF 	  i_ifDrive.etAxisState <> MOIN.ET_AxisState.Disabled
		  AND i_ifDrive.etAxisState <> MOIN.ET_AxisState.ErrorStop
		  AND i_ifDrive.etAxisState <> MOIN.ET_AxisState.Standstill
		  AND i_ifDrive.etAxisState <> MOIN.ET_AxisState.Stopping
		THEN
			fbStop.Execute 			:= TRUE;
			fbStop.Deceleration 	:= i_ifDrive.lrErrorStopDec;
			fbStop.Jerk 			:= i_ifDrive.lrErrorStopJerk;
		END_IF

		fbStop();

		//stopping done
		IF 	  i_ifDrive.etAxisState = MOIN.ET_AxisState.Disabled
		  OR  i_ifDrive.etAxisState = MOIN.ET_AxisState.ErrorStop
		  OR  i_ifDrive.etAxisState = MOIN.ET_AxisState.Standstill
		  OR  fbStop.Done
		THEN
			xInterfacesInitialised := FALSE;
			fbStop( Axis := i_ifDrive, Execute := FALSE );
			q_xInPosition	:= FALSE;
			q_xActive		:= FALSE;
			q_xReady		:= FALSE;
			SetDiagOutput(	i_etDiag	:= GD.ET_Diag.OK,
							i_etDiagExt := PDL_ET_DiagExt.Disabled,
							i_sMsg		:= '');

			diState			:= 0;
		END_IF

		//error
		IF fbStop.Error AND fbStop.ErrorId <> PLCO.ET_Result.StoppingInterrupted THEN
			q_xMotionInstructionActive	:= FALSE;

			SetDiagOutput(	i_etDiag	:= GD.ET_Diag.UnexpectedProgramBehavior,
							i_etDiagExt := PDL_ET_DiagExt.UnexpectedFeedback,
							i_sMsg		:= CONCAT('MC_Stop.ErrorID: ', PLCO.FC_EtResultToString( fbStop.ErrorID ) ));
			fbStop( Execute := FALSE );
		END_IF
{endregion}

END_CASE
(*--------------------------------------------------------------------------------------------------------------------------------------------*)
